(* Logix 5000 project; controller NWGG 1756-L72 rev 35.12; software revision 35.00; part 7 of 19 *)
(* tags used below, declared in another part *)
   _11_BINDICA : ALIAS FOR B15[11].0;
   _11_BINDICA1 : ALIAS FOR B15[11].1;
   _11_GATE_PO : ALIAS FOR I16[0];
   _11_GATE_PO1 : ALIAS FOR N14[11];
   _12_BINDICA : ALIAS FOR B15[12].0;
   _12_BINDICA1 : ALIAS FOR B15[12].1;
   _12_GATE_PO : ALIAS FOR I16[1];
   _12_GATE_PO1 : ALIAS FOR N14[12];
   _13_BINDICA : ALIAS FOR B15[13].0;
   _13_BINDICA1 : ALIAS FOR B15[13].1;
   _13_GATE_PO : ALIAS FOR I16[2];
   _13_GATE_PO1 : ALIAS FOR N14[13];
   _14_BINDICA : ALIAS FOR B15[14].0;
   _14_BINDICA1 : ALIAS FOR B15[14].1;
   _14_GATE_PO : ALIAS FOR I16[3];
   _14_GATE_PO1 : ALIAS FOR N14[14];
   _15_BINDICA : ALIAS FOR B15[15].0;
   _15_BINDICA1 : ALIAS FOR B15[15].1;
   _15_GATE_PO : ALIAS FOR I16[4];
   _15_GATE_PO1 : ALIAS FOR N14[15];
   _16_BINDICA : ALIAS FOR B15[16].0;
   _16_BINDICA1 : ALIAS FOR B15[16].1;
   _16_GATE_PO : ALIAS FOR I16[5];
   _16_GATE_PO1 : ALIAS FOR N14[16];
   _17_BINDICA : ALIAS FOR B15[17].0;
   _17_BINDICA1 : ALIAS FOR B15[17].1;
   _17_GATE_PO : ALIAS FOR I16[6];
   _17_GATE_PO1 : ALIAS FOR N14[17];
   _21_BINDICA : ALIAS FOR B15[21].0;
   _21_BINDICA1 : ALIAS FOR B15[21].1;
   _21_GATE_PO : ALIAS FOR I16[7];
   _21_GATE_PO1 : ALIAS FOR N14[21];
   _22_BINDICA : ALIAS FOR B15[22].0;
   _22_BINDICA1 : ALIAS FOR B15[22].1;
   _22_GATE_PO : ALIAS FOR I17[0];
   _22_GATE_PO1 : ALIAS FOR N14[22];
   _23_BINDICA : ALIAS FOR B15[23].0;
   _23_BINDICA1 : ALIAS FOR B15[23].1;
   _23_GATE_PO : ALIAS FOR I17[1];
   _23_GATE_PO1 : ALIAS FOR N14[23];
   _24_BINDICA : ALIAS FOR B15[24].0;
   _24_BINDICA1 : ALIAS FOR B15[24].1;
   _24_GATE_PO : ALIAS FOR I17[2];
   _24_GATE_PO1 : ALIAS FOR N14[24];
   _25_BINDICA : ALIAS FOR B15[25].0;
   _25_BINDICA1 : ALIAS FOR B15[25].1;
   _25_GATE_PO : ALIAS FOR I17[3];
   _25_GATE_PO1 : ALIAS FOR N14[25];
   _26_BINDICA : ALIAS FOR B15[26].0;
   _26_BINDICA1 : ALIAS FOR B15[26].1;
   _26_GATE_PO : ALIAS FOR I17[4];
   _26_GATE_PO1 : ALIAS FOR N14[26];
   _41_GATE_PO : ALIAS FOR I18[0];
   _41_GATE_PO1 : ALIAS FOR N14[41];
   _42_GATE_PO : ALIAS FOR I18[1];
   _42_GATE_PO1 : ALIAS FOR N14[42];
   _700_AIR_GA : ALIAS FOR I8.3;
   _701_AIR_GA : ALIAS FOR I8.5;
   _708G_BIN_1 : ALIAS FOR O9.15;
   _709G_BIN_1 : ALIAS FOR O10.15;
   A_HOLD_REL : ALIAS FOR B3[1].5;
   A_STPB_AUT : ALIAS FOR B3[1].1;
   Analog : AI[160];
   CAL_K_FACT : ALIAS FOR F8[0];
   CAL_RESET : ALIAS FOR B15[50].0;
   CIMBRA_BIN : ALIAS FOR I25[3].10;
   CIMBRIA_BI : ALIAS FOR B15[30].0;
   CIMBRIA_BI1 : ALIAS FOR B15[30].1;
   CIMBRIA_HI : ALIAS FOR B15[30].2;
   CONC13_PUM : ALIAS FOR N7[83];
   CONC19_PUM : ALIAS FOR N7[89];
   CONC_13_NO : ALIAS FOR B21[8].15;
   CONC_19_NO : ALIAS FOR B21[9].15;
   I1_000_Bit00 : ALIAS FOR I1.0;
   I1_000_Bit01 : ALIAS FOR I1.1;
   I1_000_Bit03 : ALIAS FOR I1.3;
   I1_000_Bit04 : ALIAS FOR I1.4;
   I1_000_Bit06 : ALIAS FOR I1.6;
   I1_000_Bit07 : ALIAS FOR I1.7;
   I1_000_Bit09 : ALIAS FOR I1.9;
   I1_000_Bit10 : ALIAS FOR I1.10;
   I1_000_Bit12 : ALIAS FOR I1.12;
   I1_000_Bit13 : ALIAS FOR I1.13;
   I1_000_Bit15 : ALIAS FOR I1.15;
   I24_021_Bit00 : ALIAS FOR I24[21].0;
   I24_021_Bit01 : ALIAS FOR I24[21].1;
   I24_021_Bit02 : ALIAS FOR I24[21].2;
   I2_000_Bit00 : ALIAS FOR I2.0;
   I2_000_Bit03 : ALIAS FOR I2.3;
   I2_000_Bit06 : ALIAS FOR I2.6;
   I2_000_Bit09 : ALIAS FOR I2.9;
   I2_000_Bit12 : ALIAS FOR I2.12;
   I3_000_Bit00 : ALIAS FOR I3.0;
   I3_000_Bit03 : ALIAS FOR I3.3;
   I3_000_Bit06 : ALIAS FOR I3.6;
   I4_000_Bit09 : ALIAS FOR I4.9;
   I4_000_Bit10 : ALIAS FOR I4.10;
   I4_000_Bit11 : ALIAS FOR I4.11;
   I4_000_Bit12 : ALIAS FOR I4.12;
   I4_000_Bit13 : ALIAS FOR I4.13;
   I4_000_Bit14 : ALIAS FOR I4.14;
   I4_000_Bit15 : ALIAS FOR I4.15;
   K_FACTOR : ALIAS FOR N14[80];
   P1_ALARM_N : ALIAS FOR T4[81];
   P1_ALARM_N1 : ALIAS FOR T4[82];
   P1_NO_FLOW : ALIAS FOR B12[1].3;
   P1_SEC_SEL : ALIAS FOR B17[1].1;
   P2_ALARM_N : ALIAS FOR T4[83];
   P2_ALARM_N1 : ALIAS FOR T4[84];
   P2_NO_FLOW : ALIAS FOR B12[2].3;
   P2_SEC_SEL : ALIAS FOR B17[1].2;
   P3_ALARM_N : ALIAS FOR T4[85];
   P3_ALARM_N1 : ALIAS FOR T4[86];
   P3_NO_FLOW : ALIAS FOR B12[3].3;
   P3_SEC_SEL : ALIAS FOR B17[1].3;
   P4_SEC_SEL : ALIAS FOR B17[1].4;
   T11_CAL_CL : ALIAS FOR B15[51].3;
   T11_CAL_LA : ALIAS FOR B15[51].2;
   T11_CAL_OP : ALIAS FOR B15[51].4;
   T11_CAL_ST : ALIAS FOR B15[51].1;
   T11_CORREC : ALIAS FOR F8[2];
   T11_K_FACT : ALIAS FOR F8[1];
   T11_LOW_BI : ALIAS FOR B15[11].2;
   T11_NO_PAS : ALIAS FOR B17[11].2;
   T12_CAL_CL : ALIAS FOR B15[52].3;
   T12_CAL_LA : ALIAS FOR B15[52].2;
   T12_CAL_OP : ALIAS FOR B15[52].4;
   T12_CAL_ST : ALIAS FOR B15[52].1;
   T12_CORREC : ALIAS FOR F8[4];
   T12_K_FACT : ALIAS FOR F8[3];
   T12_LOW_BI : ALIAS FOR B15[12].2;
   T12_NO_PAS : ALIAS FOR B17[12].2;
   T13_CAL_CL : ALIAS FOR B15[53].3;
   T13_CAL_LA : ALIAS FOR B15[53].2;
   T13_CAL_OP : ALIAS FOR B15[53].4;
   T13_CAL_ST : ALIAS FOR B15[53].1;
   T13_CORREC : ALIAS FOR F8[6];
   T13_K_FACT : ALIAS FOR F8[5];
   T13_LOW_BI : ALIAS FOR B15[13].2;
   T13_NO_PAS : ALIAS FOR B17[13].2;
   T14_CAL_CL : ALIAS FOR B15[54].3;
   T14_CAL_LA : ALIAS FOR B15[54].2;
   T14_CAL_OP : ALIAS FOR B15[54].4;
   T14_CAL_ST : ALIAS FOR B15[54].1;
   T14_CORREC : ALIAS FOR F8[8];
   T14_K_FACT : ALIAS FOR F8[7];
   T14_LOW_BI : ALIAS FOR B15[14].2;
   T14_NO_PAS : ALIAS FOR B17[14].2;
   T15_CAL_CL : ALIAS FOR B15[55].3;
   T15_CAL_LA : ALIAS FOR B15[55].2;
   T15_CAL_OP : ALIAS FOR B15[55].4;
   T15_CAL_ST : ALIAS FOR B15[55].1;
   T15_CORREC : ALIAS FOR F8[10];
   T15_K_FACT : ALIAS FOR F8[9];
   T15_LOW_BI : ALIAS FOR B15[15].2;
   T15_NO_PAS : ALIAS FOR B17[15].2;
   T16_CAL_CL : ALIAS FOR B15[56].3;
   T16_CAL_LA : ALIAS FOR B15[56].2;
   T16_CAL_OP : ALIAS FOR B15[56].4;
   T16_CAL_ST : ALIAS FOR B15[56].1;
   T16_CORREC : ALIAS FOR F8[12];
   T16_K_FACT : ALIAS FOR F8[11];
   T16_LOW_BI : ALIAS FOR B15[16].2;
   T16_NO_PAS : ALIAS FOR B17[16].2;
   T17_CAL_CL : ALIAS FOR B15[57].3;
   T17_CAL_LA : ALIAS FOR B15[57].2;
   T17_CAL_OP : ALIAS FOR B15[57].4;
   T17_CAL_ST : ALIAS FOR B15[57].1;
   T17_CORREC : ALIAS FOR F8[14];
   T17_K_FACT : ALIAS FOR F8[13];
   T17_LOW_BI : ALIAS FOR B15[17].2;
   T17_NO_PAS : ALIAS FOR B17[17].2;
   T21_CAL_CL : ALIAS FOR B15[61].3;
   T21_CAL_LA : ALIAS FOR B15[61].2;
   T21_CAL_OP : ALIAS FOR B15[61].4;
   T21_CAL_ST : ALIAS FOR B15[61].1;
   T21_CORREC : ALIAS FOR F8[16];
   T21_K_FACT : ALIAS FOR F8[15];
   T21_LOW_BI : ALIAS FOR B15[21].2;
   T21_NO_PAS : ALIAS FOR B17[21].2;
   T22_CAL_CL : ALIAS FOR B15[62].3;
   T22_CAL_LA : ALIAS FOR B15[62].2;
   T22_CAL_OP : ALIAS FOR B15[62].4;
   T22_CAL_ST : ALIAS FOR B15[62].1;
   T22_CORREC : ALIAS FOR F8[18];
   T22_K_FACT : ALIAS FOR F8[17];
   T22_LOW_BI : ALIAS FOR B15[22].2;
   T22_NO_PAS : ALIAS FOR B17[22].2;
   T23_CAL_CL : ALIAS FOR B15[63].3;
   T23_CAL_LA : ALIAS FOR B15[63].2;
   T23_CAL_OP : ALIAS FOR B15[63].4;
   T23_CAL_ST : ALIAS FOR B15[63].1;
   T23_CORREC : ALIAS FOR F8[20];
   T23_K_FACT : ALIAS FOR F8[19];
   T23_LOW_BI : ALIAS FOR B15[23].2;
   T23_NO_PAS : ALIAS FOR B17[23].2;
   T24_CAL_CL : ALIAS FOR B15[64].3;
   T24_CAL_LA : ALIAS FOR B15[64].2;
   T24_CAL_OP : ALIAS FOR B15[64].4;
   T24_CAL_ST : ALIAS FOR B15[64].1;
   T24_CORREC : ALIAS FOR F8[22];
   T24_K_FACT : ALIAS FOR F8[21];
   T24_LOW_BI : ALIAS FOR B15[24].2;
   T24_NO_PAS : ALIAS FOR B17[24].2;
   T25_CAL_CL : ALIAS FOR B15[65].3;
   T25_CAL_LA : ALIAS FOR B15[65].2;
   T25_CAL_OP : ALIAS FOR B15[65].4;
   T25_CAL_ST : ALIAS FOR B15[65].1;
   T25_CORREC : ALIAS FOR F8[24];
   T25_K_FACT : ALIAS FOR F8[23];
   T25_LOW_BI : ALIAS FOR B15[25].2;
   T25_NO_PAS : ALIAS FOR B17[25].2;
   T26_CAL_CL : ALIAS FOR B15[66].3;
   T26_CAL_LA : ALIAS FOR B15[66].2;
   T26_CAL_OP : ALIAS FOR B15[66].4;
   T26_CAL_ST : ALIAS FOR B15[66].1;
   T26_CORREC : ALIAS FOR F8[26];
   T26_K_FACT : ALIAS FOR F8[25];
   T26_LOW_BI : ALIAS FOR B15[26].2;
   T26_NO_PAS : ALIAS FOR B17[26].2;
   TK11_PUMP : ALIAS FOR N7[70];
   TK12_PUMP : ALIAS FOR N7[71];
   TK13_PUMP : ALIAS FOR N7[72];
   TK14_PUMP : ALIAS FOR N7[73];
   TK15_PUMP : ALIAS FOR N7[74];
   TK16_PUMP : ALIAS FOR N7[75];
   TK17_PUMP : ALIAS FOR N7[76];
   TK21_PUMP : ALIAS FOR N7[77];
   TK22_PUMP : ALIAS FOR N7[78];
   TK23_PUMP : ALIAS FOR N7[79];
   TK24_PUMP : ALIAS FOR N7[80];
   TK25_PUMP : ALIAS FOR N7[81];
   TK26_PUMP : ALIAS FOR N7[82];
(* _2_MAIN, continued *)

ROUTINE _37_BINDICATOR   (* ladder *)
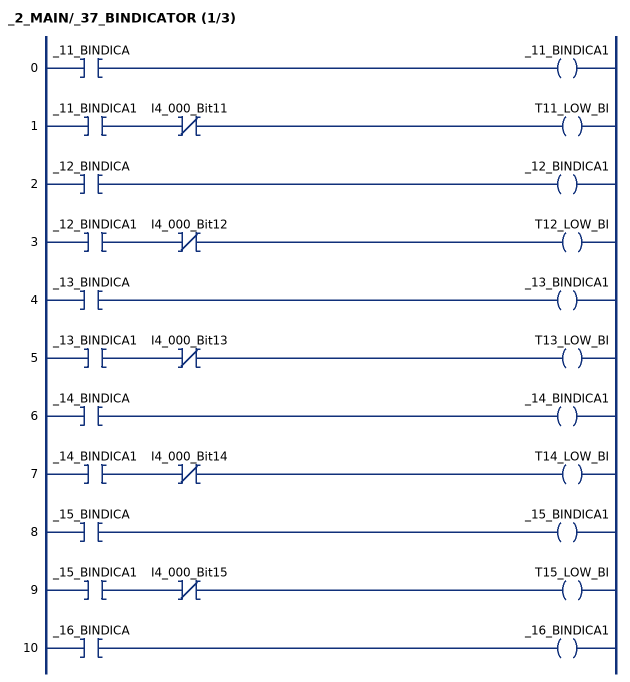
   0: XIC(_11_BINDICA)OTE(_11_BINDICA1);
   1: XIC(_11_BINDICA1)XIO(I4_000_Bit11)OTE(T11_LOW_BI);
   2: XIC(_12_BINDICA)OTE(_12_BINDICA1);
   3: XIC(_12_BINDICA1)XIO(I4_000_Bit12)OTE(T12_LOW_BI);
   4: XIC(_13_BINDICA)OTE(_13_BINDICA1);
   5: XIC(_13_BINDICA1)XIO(I4_000_Bit13)OTE(T13_LOW_BI);
   6: XIC(_14_BINDICA)OTE(_14_BINDICA1);
   7: XIC(_14_BINDICA1)XIO(I4_000_Bit14)OTE(T14_LOW_BI);
   8: XIC(_15_BINDICA)OTE(_15_BINDICA1);
   9: XIC(_15_BINDICA1)XIO(I4_000_Bit15)OTE(T15_LOW_BI);
   10: XIC(_16_BINDICA)OTE(_16_BINDICA1);
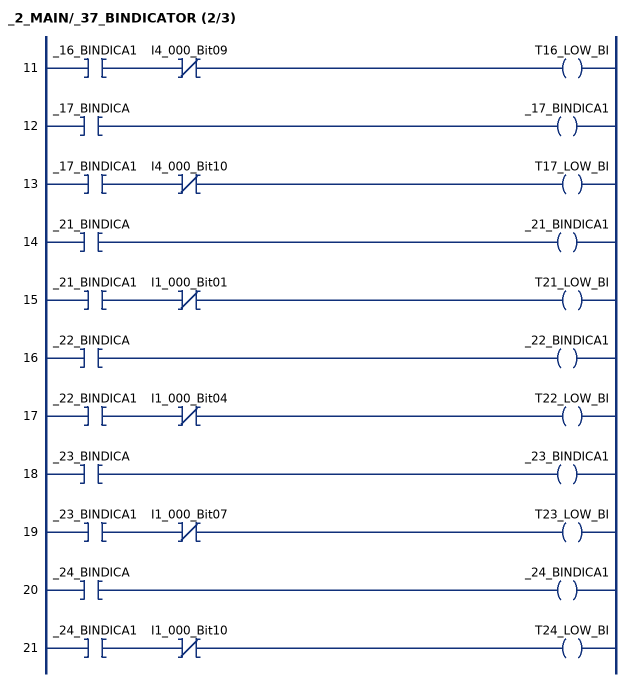
   11: XIC(_16_BINDICA1)XIO(I4_000_Bit09)OTE(T16_LOW_BI);
   12: XIC(_17_BINDICA)OTE(_17_BINDICA1);
   13: XIC(_17_BINDICA1)XIO(I4_000_Bit10)OTE(T17_LOW_BI);
   14: XIC(_21_BINDICA)OTE(_21_BINDICA1);
   15: XIC(_21_BINDICA1)XIO(I1_000_Bit01)OTE(T21_LOW_BI);
   16: XIC(_22_BINDICA)OTE(_22_BINDICA1);
   17: XIC(_22_BINDICA1)XIO(I1_000_Bit04)OTE(T22_LOW_BI);
   18: XIC(_23_BINDICA)OTE(_23_BINDICA1);
   19: XIC(_23_BINDICA1)XIO(I1_000_Bit07)OTE(T23_LOW_BI);
   20: XIC(_24_BINDICA)OTE(_24_BINDICA1);
   21: XIC(_24_BINDICA1)XIO(I1_000_Bit10)OTE(T24_LOW_BI);
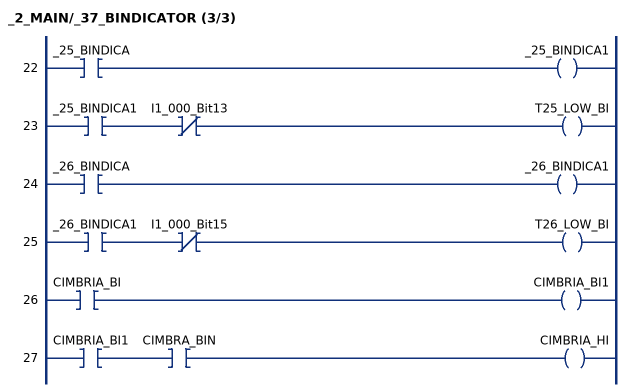
   22: XIC(_25_BINDICA)OTE(_25_BINDICA1);
   23: XIC(_25_BINDICA1)XIO(I1_000_Bit13)OTE(T25_LOW_BI);
   24: XIC(_26_BINDICA)OTE(_26_BINDICA1);
   25: XIC(_26_BINDICA1)XIO(I1_000_Bit15)OTE(T26_LOW_BI);
   26: XIC(CIMBRIA_BI)OTE(CIMBRIA_BI1);
   27: XIC(CIMBRIA_BI1)XIC(CIMBRA_BIN)OTE(CIMBRIA_HI);
END_ROUTINE

ROUTINE _38_GATE_ADJST   (* ladder *)
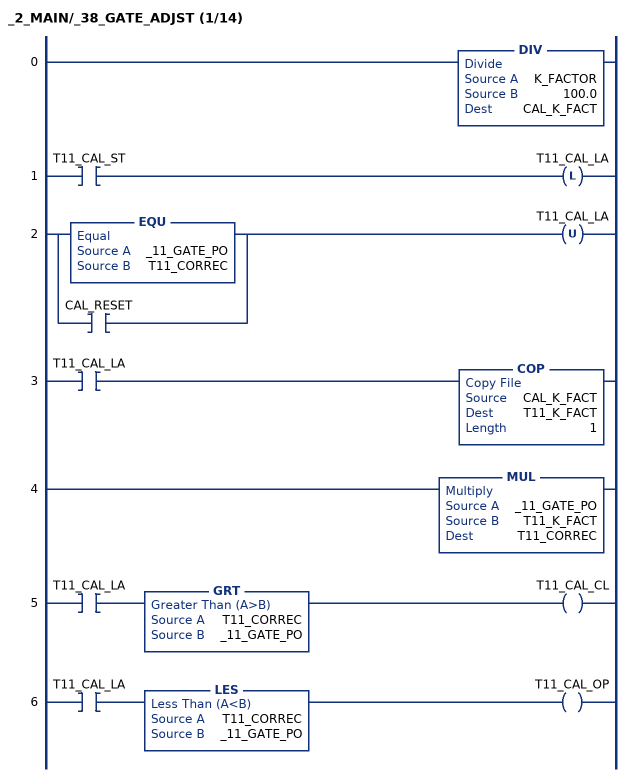
   0: DIV(K_FACTOR,100.0,CAL_K_FACT);
   1: XIC(T11_CAL_ST)OTL(T11_CAL_LA);
   2: [EQU(_11_GATE_PO,T11_CORREC) ,XIC(CAL_RESET) ]OTU(T11_CAL_LA);
   3: XIC(T11_CAL_LA)COP(CAL_K_FACT,T11_K_FACT,1);
   4: MUL(_11_GATE_PO,T11_K_FACT,T11_CORREC);
   5: XIC(T11_CAL_LA)GRT(T11_CORREC,_11_GATE_PO)OTE(T11_CAL_CL);
   6: XIC(T11_CAL_LA)LES(T11_CORREC,_11_GATE_PO)OTE(T11_CAL_OP);
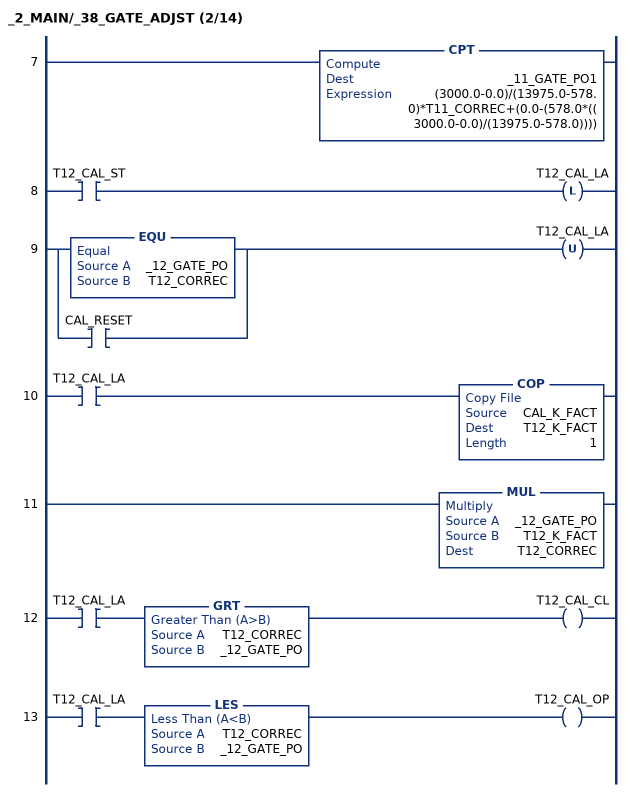
   7: CPT(_11_GATE_PO1,(3000.0-0.0)/(13975.0-578.0)*T11_CORREC+(0.0-(578.0*((3000.0-0.0)/(13975.0-578.0)))));
   8: XIC(T12_CAL_ST)OTL(T12_CAL_LA);
   9: [EQU(_12_GATE_PO,T12_CORREC) ,XIC(CAL_RESET) ]OTU(T12_CAL_LA);
   10: XIC(T12_CAL_LA)COP(CAL_K_FACT,T12_K_FACT,1);
   11: MUL(_12_GATE_PO,T12_K_FACT,T12_CORREC);
   12: XIC(T12_CAL_LA)GRT(T12_CORREC,_12_GATE_PO)OTE(T12_CAL_CL);
   13: XIC(T12_CAL_LA)LES(T12_CORREC,_12_GATE_PO)OTE(T12_CAL_OP);
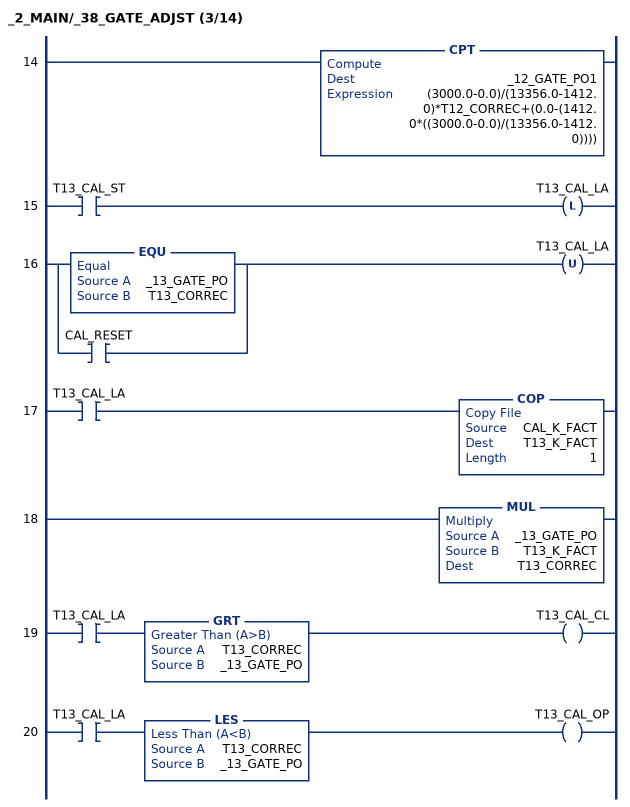
   14: CPT(_12_GATE_PO1,(3000.0-0.0)/(13356.0-1412.0)*T12_CORREC+(0.0-(1412.0*((3000.0-0.0)/(13356.0-1412.0)))));
   15: XIC(T13_CAL_ST)OTL(T13_CAL_LA);
   16: [EQU(_13_GATE_PO,T13_CORREC) ,XIC(CAL_RESET) ]OTU(T13_CAL_LA);
   17: XIC(T13_CAL_LA)COP(CAL_K_FACT,T13_K_FACT,1);
   18: MUL(_13_GATE_PO,T13_K_FACT,T13_CORREC);
   19: XIC(T13_CAL_LA)GRT(T13_CORREC,_13_GATE_PO)OTE(T13_CAL_CL);
   20: XIC(T13_CAL_LA)LES(T13_CORREC,_13_GATE_PO)OTE(T13_CAL_OP);
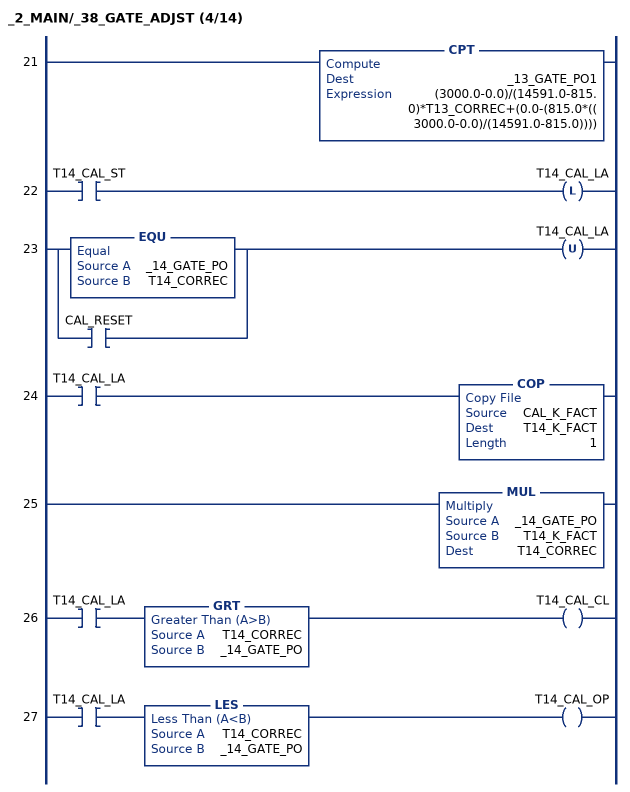
   21: CPT(_13_GATE_PO1,(3000.0-0.0)/(14591.0-815.0)*T13_CORREC+(0.0-(815.0*((3000.0-0.0)/(14591.0-815.0)))));
   22: XIC(T14_CAL_ST)OTL(T14_CAL_LA);
   23: [EQU(_14_GATE_PO,T14_CORREC) ,XIC(CAL_RESET) ]OTU(T14_CAL_LA);
   24: XIC(T14_CAL_LA)COP(CAL_K_FACT,T14_K_FACT,1);
   25: MUL(_14_GATE_PO,T14_K_FACT,T14_CORREC);
   26: XIC(T14_CAL_LA)GRT(T14_CORREC,_14_GATE_PO)OTE(T14_CAL_CL);
   27: XIC(T14_CAL_LA)LES(T14_CORREC,_14_GATE_PO)OTE(T14_CAL_OP);
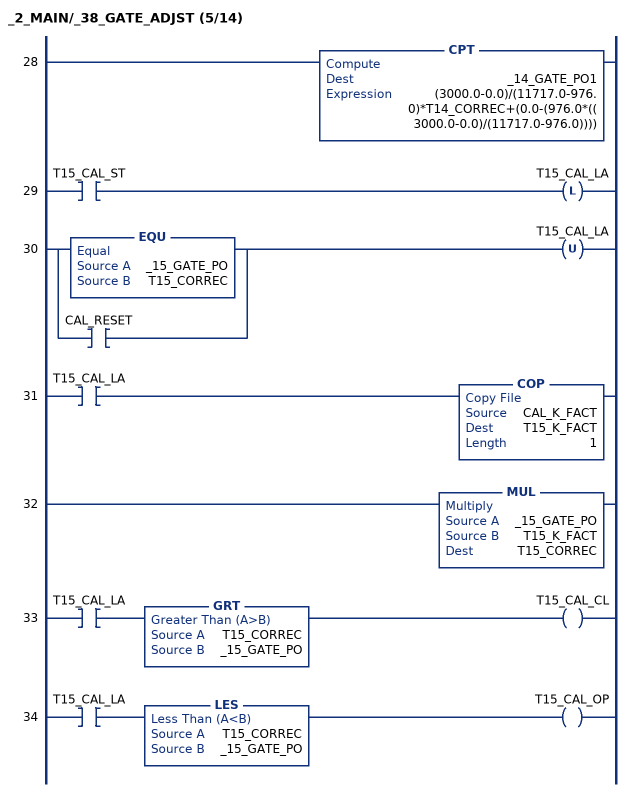
   28: CPT(_14_GATE_PO1,(3000.0-0.0)/(11717.0-976.0)*T14_CORREC+(0.0-(976.0*((3000.0-0.0)/(11717.0-976.0)))));
   29: XIC(T15_CAL_ST)OTL(T15_CAL_LA);
   30: [EQU(_15_GATE_PO,T15_CORREC) ,XIC(CAL_RESET) ]OTU(T15_CAL_LA);
   31: XIC(T15_CAL_LA)COP(CAL_K_FACT,T15_K_FACT,1);
   32: MUL(_15_GATE_PO,T15_K_FACT,T15_CORREC);
   33: XIC(T15_CAL_LA)GRT(T15_CORREC,_15_GATE_PO)OTE(T15_CAL_CL);
   34: XIC(T15_CAL_LA)LES(T15_CORREC,_15_GATE_PO)OTE(T15_CAL_OP);
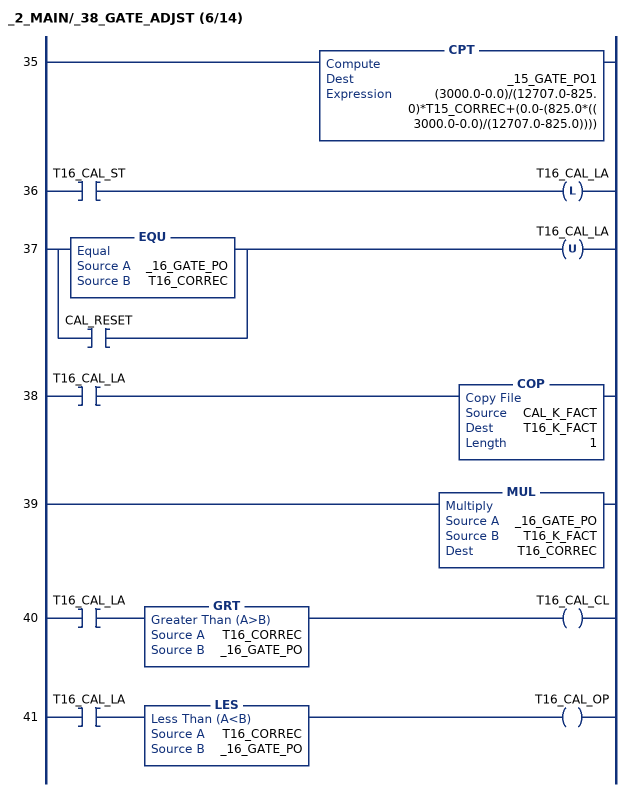
   35: CPT(_15_GATE_PO1,(3000.0-0.0)/(12707.0-825.0)*T15_CORREC+(0.0-(825.0*((3000.0-0.0)/(12707.0-825.0)))));
   36: XIC(T16_CAL_ST)OTL(T16_CAL_LA);
   37: [EQU(_16_GATE_PO,T16_CORREC) ,XIC(CAL_RESET) ]OTU(T16_CAL_LA);
   38: XIC(T16_CAL_LA)COP(CAL_K_FACT,T16_K_FACT,1);
   39: MUL(_16_GATE_PO,T16_K_FACT,T16_CORREC);
   40: XIC(T16_CAL_LA)GRT(T16_CORREC,_16_GATE_PO)OTE(T16_CAL_CL);
   41: XIC(T16_CAL_LA)LES(T16_CORREC,_16_GATE_PO)OTE(T16_CAL_OP);
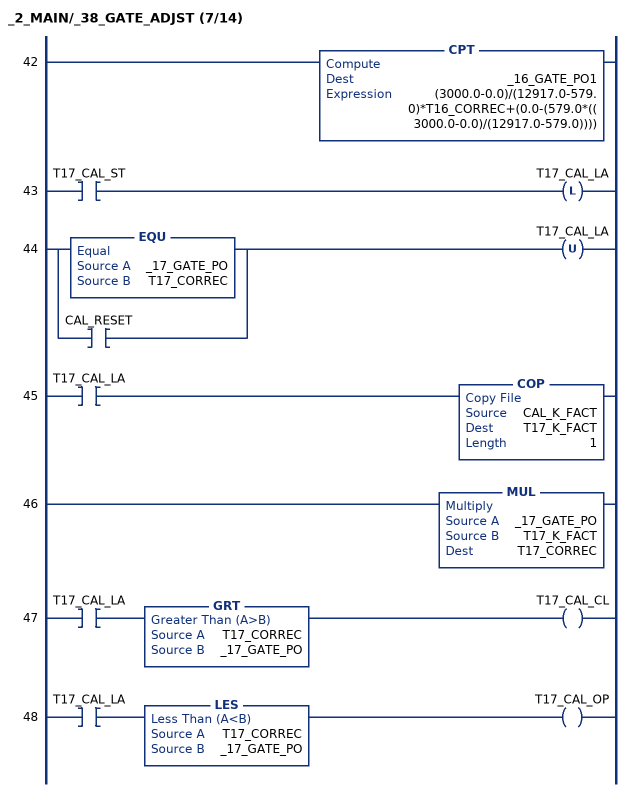
   42: CPT(_16_GATE_PO1,(3000.0-0.0)/(12917.0-579.0)*T16_CORREC+(0.0-(579.0*((3000.0-0.0)/(12917.0-579.0)))));
   43: XIC(T17_CAL_ST)OTL(T17_CAL_LA);
   44: [EQU(_17_GATE_PO,T17_CORREC) ,XIC(CAL_RESET) ]OTU(T17_CAL_LA);
   45: XIC(T17_CAL_LA)COP(CAL_K_FACT,T17_K_FACT,1);
   46: MUL(_17_GATE_PO,T17_K_FACT,T17_CORREC);
   47: XIC(T17_CAL_LA)GRT(T17_CORREC,_17_GATE_PO)OTE(T17_CAL_CL);
   48: XIC(T17_CAL_LA)LES(T17_CORREC,_17_GATE_PO)OTE(T17_CAL_OP);
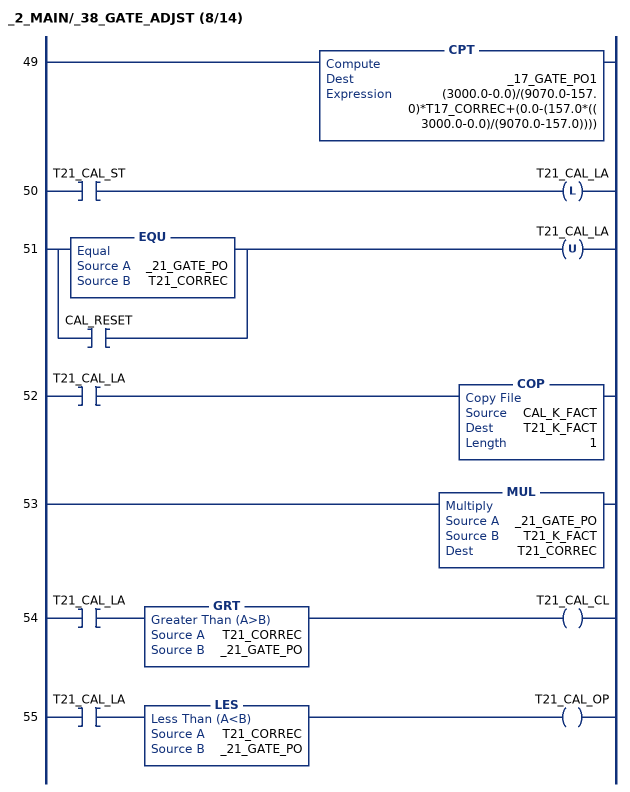
   49: CPT(_17_GATE_PO1,(3000.0-0.0)/(9070.0-157.0)*T17_CORREC+(0.0-(157.0*((3000.0-0.0)/(9070.0-157.0)))));
   50: XIC(T21_CAL_ST)OTL(T21_CAL_LA);
   51: [EQU(_21_GATE_PO,T21_CORREC) ,XIC(CAL_RESET) ]OTU(T21_CAL_LA);
   52: XIC(T21_CAL_LA)COP(CAL_K_FACT,T21_K_FACT,1);
   53: MUL(_21_GATE_PO,T21_K_FACT,T21_CORREC);
   54: XIC(T21_CAL_LA)GRT(T21_CORREC,_21_GATE_PO)OTE(T21_CAL_CL);
   55: XIC(T21_CAL_LA)LES(T21_CORREC,_21_GATE_PO)OTE(T21_CAL_OP);
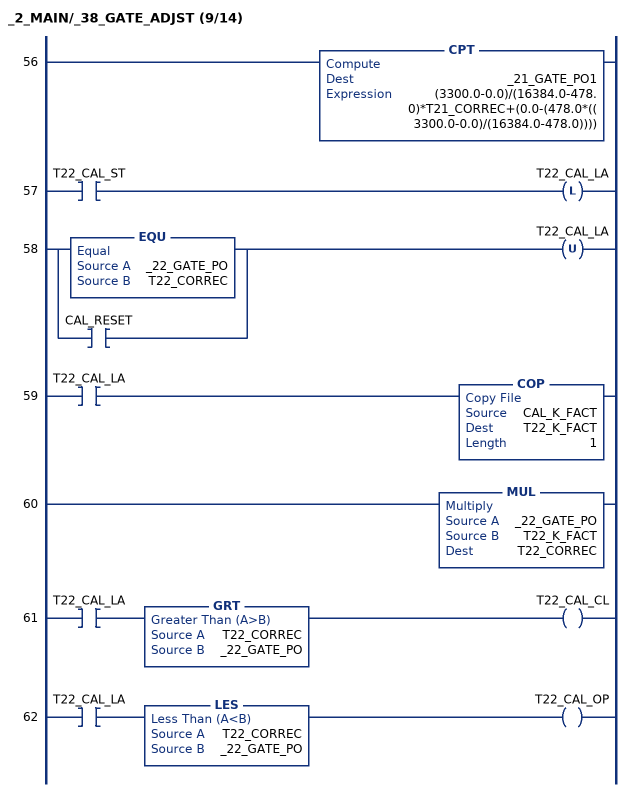
   56: CPT(_21_GATE_PO1,(3300.0-0.0)/(16384.0-478.0)*T21_CORREC+(0.0-(478.0*((3300.0-0.0)/(16384.0-478.0)))));
   57: XIC(T22_CAL_ST)OTL(T22_CAL_LA);
   58: [EQU(_22_GATE_PO,T22_CORREC) ,XIC(CAL_RESET) ]OTU(T22_CAL_LA);
   59: XIC(T22_CAL_LA)COP(CAL_K_FACT,T22_K_FACT,1);
   60: MUL(_22_GATE_PO,T22_K_FACT,T22_CORREC);
   61: XIC(T22_CAL_LA)GRT(T22_CORREC,_22_GATE_PO)OTE(T22_CAL_CL);
   62: XIC(T22_CAL_LA)LES(T22_CORREC,_22_GATE_PO)OTE(T22_CAL_OP);
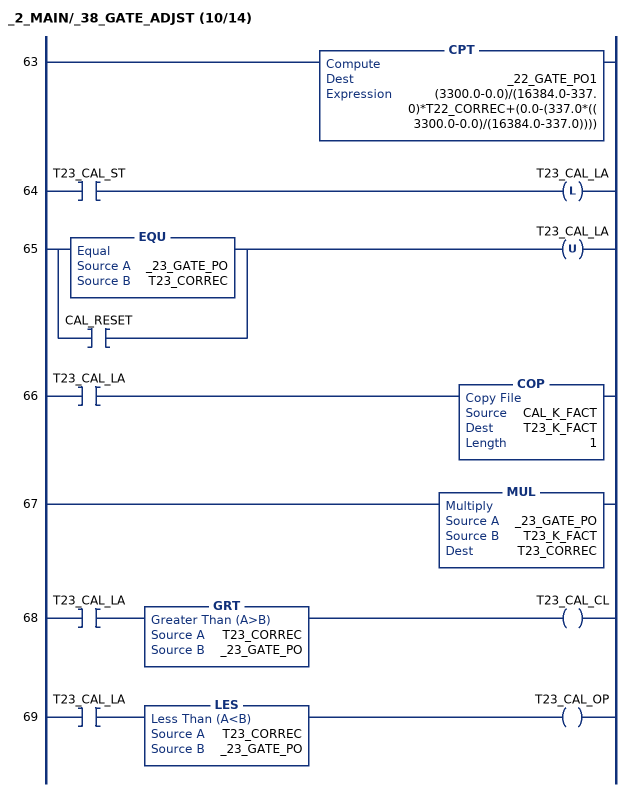
   63: CPT(_22_GATE_PO1,(3300.0-0.0)/(16384.0-337.0)*T22_CORREC+(0.0-(337.0*((3300.0-0.0)/(16384.0-337.0)))));
   64: XIC(T23_CAL_ST)OTL(T23_CAL_LA);
   65: [EQU(_23_GATE_PO,T23_CORREC) ,XIC(CAL_RESET) ]OTU(T23_CAL_LA);
   66: XIC(T23_CAL_LA)COP(CAL_K_FACT,T23_K_FACT,1);
   67: MUL(_23_GATE_PO,T23_K_FACT,T23_CORREC);
   68: XIC(T23_CAL_LA)GRT(T23_CORREC,_23_GATE_PO)OTE(T23_CAL_CL);
   69: XIC(T23_CAL_LA)LES(T23_CORREC,_23_GATE_PO)OTE(T23_CAL_OP);
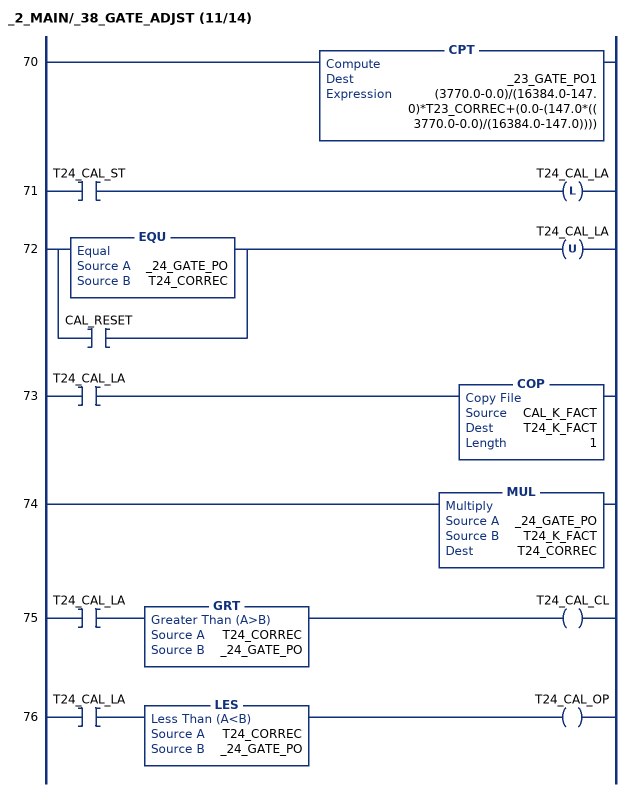
   70: CPT(_23_GATE_PO1,(3770.0-0.0)/(16384.0-147.0)*T23_CORREC+(0.0-(147.0*((3770.0-0.0)/(16384.0-147.0)))));
   71: XIC(T24_CAL_ST)OTL(T24_CAL_LA);
   72: [EQU(_24_GATE_PO,T24_CORREC) ,XIC(CAL_RESET) ]OTU(T24_CAL_LA);
   73: XIC(T24_CAL_LA)COP(CAL_K_FACT,T24_K_FACT,1);
   74: MUL(_24_GATE_PO,T24_K_FACT,T24_CORREC);
   75: XIC(T24_CAL_LA)GRT(T24_CORREC,_24_GATE_PO)OTE(T24_CAL_CL);
   76: XIC(T24_CAL_LA)LES(T24_CORREC,_24_GATE_PO)OTE(T24_CAL_OP);
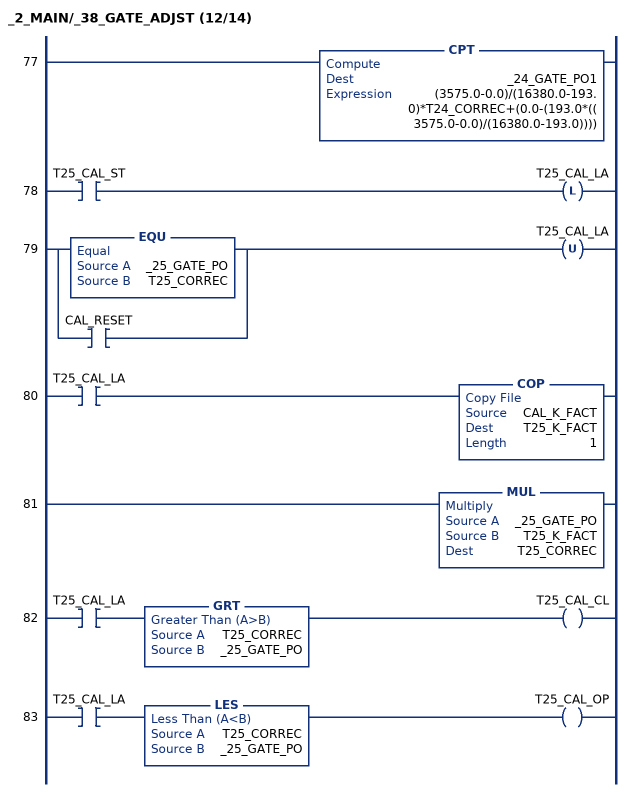
   77: CPT(_24_GATE_PO1,(3575.0-0.0)/(16380.0-193.0)*T24_CORREC+(0.0-(193.0*((3575.0-0.0)/(16380.0-193.0)))));
   78: XIC(T25_CAL_ST)OTL(T25_CAL_LA);
   79: [EQU(_25_GATE_PO,T25_CORREC) ,XIC(CAL_RESET) ]OTU(T25_CAL_LA);
   80: XIC(T25_CAL_LA)COP(CAL_K_FACT,T25_K_FACT,1);
   81: MUL(_25_GATE_PO,T25_K_FACT,T25_CORREC);
   82: XIC(T25_CAL_LA)GRT(T25_CORREC,_25_GATE_PO)OTE(T25_CAL_CL);
   83: XIC(T25_CAL_LA)LES(T25_CORREC,_25_GATE_PO)OTE(T25_CAL_OP);
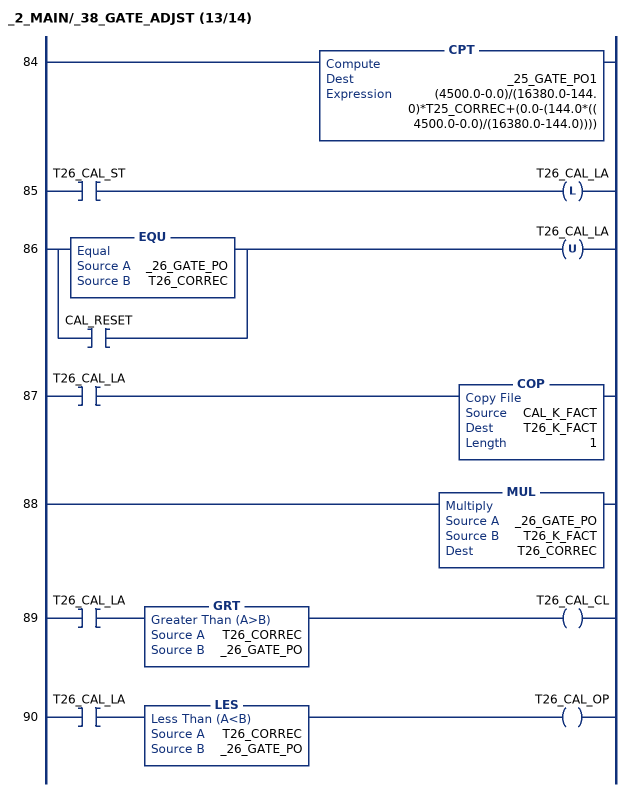
   84: CPT(_25_GATE_PO1,(4500.0-0.0)/(16380.0-144.0)*T25_CORREC+(0.0-(144.0*((4500.0-0.0)/(16380.0-144.0)))));
   85: XIC(T26_CAL_ST)OTL(T26_CAL_LA);
   86: [EQU(_26_GATE_PO,T26_CORREC) ,XIC(CAL_RESET) ]OTU(T26_CAL_LA);
   87: XIC(T26_CAL_LA)COP(CAL_K_FACT,T26_K_FACT,1);
   88: MUL(_26_GATE_PO,T26_K_FACT,T26_CORREC);
   89: XIC(T26_CAL_LA)GRT(T26_CORREC,_26_GATE_PO)OTE(T26_CAL_CL);
   90: XIC(T26_CAL_LA)LES(T26_CORREC,_26_GATE_PO)OTE(T26_CAL_OP);
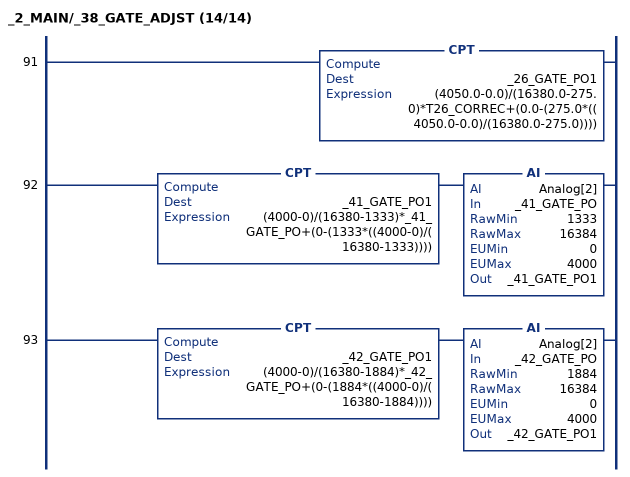
   91: CPT(_26_GATE_PO1,(4050.0-0.0)/(16380.0-275.0)*T26_CORREC+(0.0-(275.0*((4050.0-0.0)/(16380.0-275.0)))));
   92: CPT(_41_GATE_PO1,(4000-0)/(16380-1333)*_41_GATE_PO+(0-(1333*((4000-0)/(16380-1333)))))AI(Analog[2],_41_GATE_PO,1333,16384,0,4000,_41_GATE_PO1);
   93: CPT(_42_GATE_PO1,(4000-0)/(16380-1884)*_42_GATE_PO+(0-(1884*((4000-0)/(16380-1884)))))AI(Analog[2],_42_GATE_PO,1884,16384,0,4000,_42_GATE_PO1);
END_ROUTINE

ROUTINE _39_PUMP_SECUR   (* ladder *)
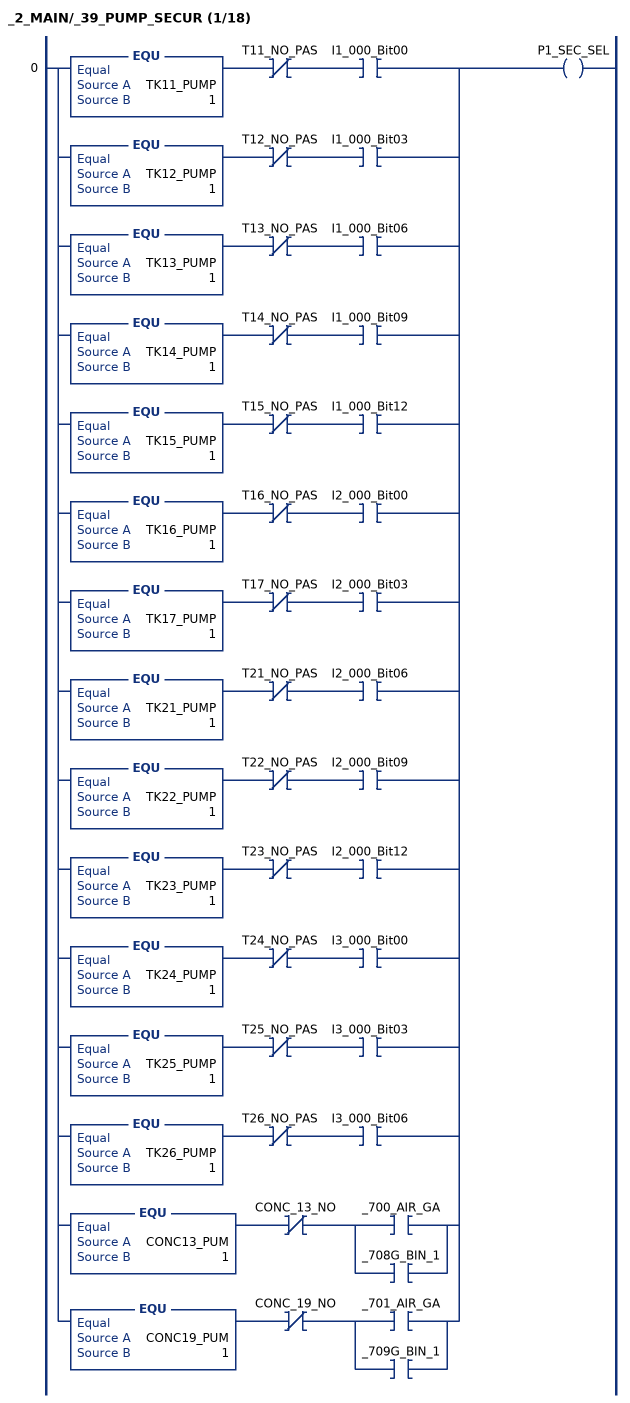
   0: [EQU(TK11_PUMP,1) XIO(T11_NO_PAS) XIC(I1_000_Bit00) ,EQU(TK12_PUMP,1) XIO(T12_NO_PAS) XIC(I1_000_Bit03) ,EQU(TK13_PUMP,1) XIO(T13_NO_PAS) XIC(I1_000_Bit06) ,EQU(TK14_PUMP,1) XIO(T14_NO_PAS) XIC(I1_000_Bit09) ,EQU(TK15_PUMP,1) XIO(T15_NO_PAS) XIC(I1_000_Bit12) ,EQU(TK16_PUMP,1) XIO(T16_NO_PAS) XIC(I2_000_Bit00) ,EQU(TK17_PUMP,1) XIO(T17_NO_PAS) XIC(I2_000_Bit03) ,EQU(TK21_PUMP,1) XIO(T21_NO_PAS) XIC(I2_000_Bit06) ,EQU(TK22_PUMP,1) XIO(T22_NO_PAS) XIC(I2_000_Bit09) ,EQU(TK23_PUMP,1) XIO(T23_NO_PAS) XIC(I2_000_Bit12) ,EQU(TK24_PUMP,1) XIO(T24_NO_PAS) XIC(I3_000_Bit00) ,EQU(TK25_PUMP,1) XIO(T25_NO_PAS) XIC(I3_000_Bit03) ,EQU(TK26_PUMP,1) XIO(T26_NO_PAS) XIC(I3_000_Bit06) ,EQU(CONC13_PUM,1) XIO(CONC_13_NO) [XIC(_700_AIR_GA) ,XIC(_708G_BIN_1) ] ,EQU(CONC19_PUM,1) XIO(CONC_19_NO) [XIC(_701_AIR_GA) ,XIC(_709G_BIN_1) ] ]OTE(P1_SEC_SEL);
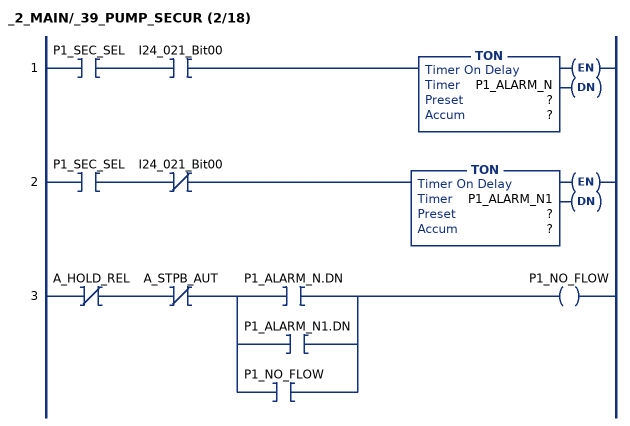
   1: XIC(P1_SEC_SEL)XIC(I24_021_Bit00)TON(P1_ALARM_N,?,?);
   2: XIC(P1_SEC_SEL)XIO(I24_021_Bit00)TON(P1_ALARM_N1,?,?);
   3: XIO(A_HOLD_REL)XIO(A_STPB_AUT)[XIC(P1_ALARM_N.DN) ,XIC(P1_ALARM_N1.DN) ,XIC(P1_NO_FLOW) ]OTE(P1_NO_FLOW);
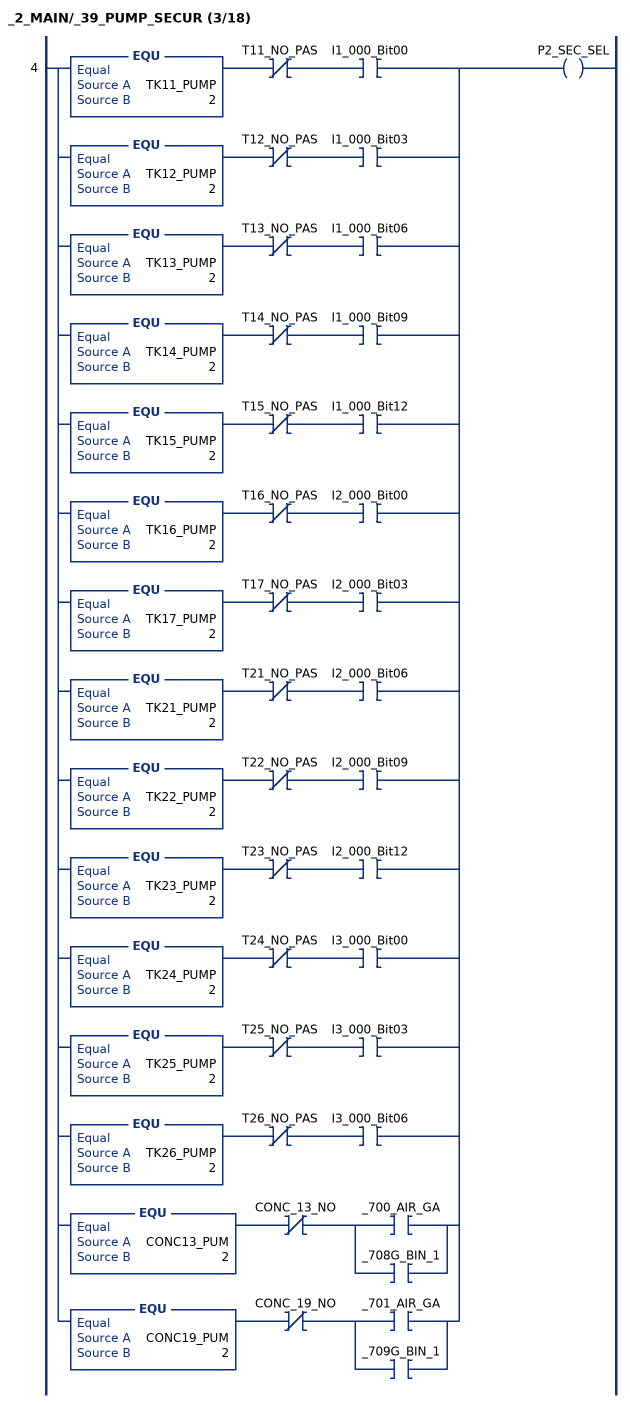
   4: [EQU(TK11_PUMP,2) XIO(T11_NO_PAS) XIC(I1_000_Bit00) ,EQU(TK12_PUMP,2) XIO(T12_NO_PAS) XIC(I1_000_Bit03) ,EQU(TK13_PUMP,2) XIO(T13_NO_PAS) XIC(I1_000_Bit06) ,EQU(TK14_PUMP,2) XIO(T14_NO_PAS) XIC(I1_000_Bit09) ,EQU(TK15_PUMP,2) XIO(T15_NO_PAS) XIC(I1_000_Bit12) ,EQU(TK16_PUMP,2) XIO(T16_NO_PAS) XIC(I2_000_Bit00) ,EQU(TK17_PUMP,2) XIO(T17_NO_PAS) XIC(I2_000_Bit03) ,EQU(TK21_PUMP,2) XIO(T21_NO_PAS) XIC(I2_000_Bit06) ,EQU(TK22_PUMP,2) XIO(T22_NO_PAS) XIC(I2_000_Bit09) ,EQU(TK23_PUMP,2) XIO(T23_NO_PAS) XIC(I2_000_Bit12) ,EQU(TK24_PUMP,2) XIO(T24_NO_PAS) XIC(I3_000_Bit00) ,EQU(TK25_PUMP,2) XIO(T25_NO_PAS) XIC(I3_000_Bit03) ,EQU(TK26_PUMP,2) XIO(T26_NO_PAS) XIC(I3_000_Bit06) ,EQU(CONC13_PUM,2) XIO(CONC_13_NO) [XIC(_700_AIR_GA) ,XIC(_708G_BIN_1) ] ,EQU(CONC19_PUM,2) XIO(CONC_19_NO) [XIC(_701_AIR_GA) ,XIC(_709G_BIN_1) ] ]OTE(P2_SEC_SEL);
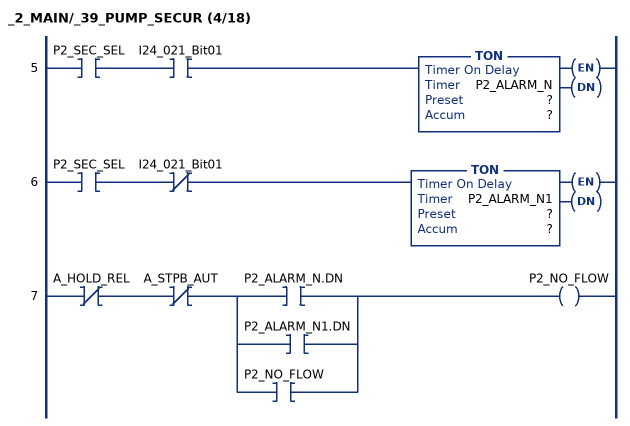
   5: XIC(P2_SEC_SEL)XIC(I24_021_Bit01)TON(P2_ALARM_N,?,?);
   6: XIC(P2_SEC_SEL)XIO(I24_021_Bit01)TON(P2_ALARM_N1,?,?);
   7: XIO(A_HOLD_REL)XIO(A_STPB_AUT)[XIC(P2_ALARM_N.DN) ,XIC(P2_ALARM_N1.DN) ,XIC(P2_NO_FLOW) ]OTE(P2_NO_FLOW);
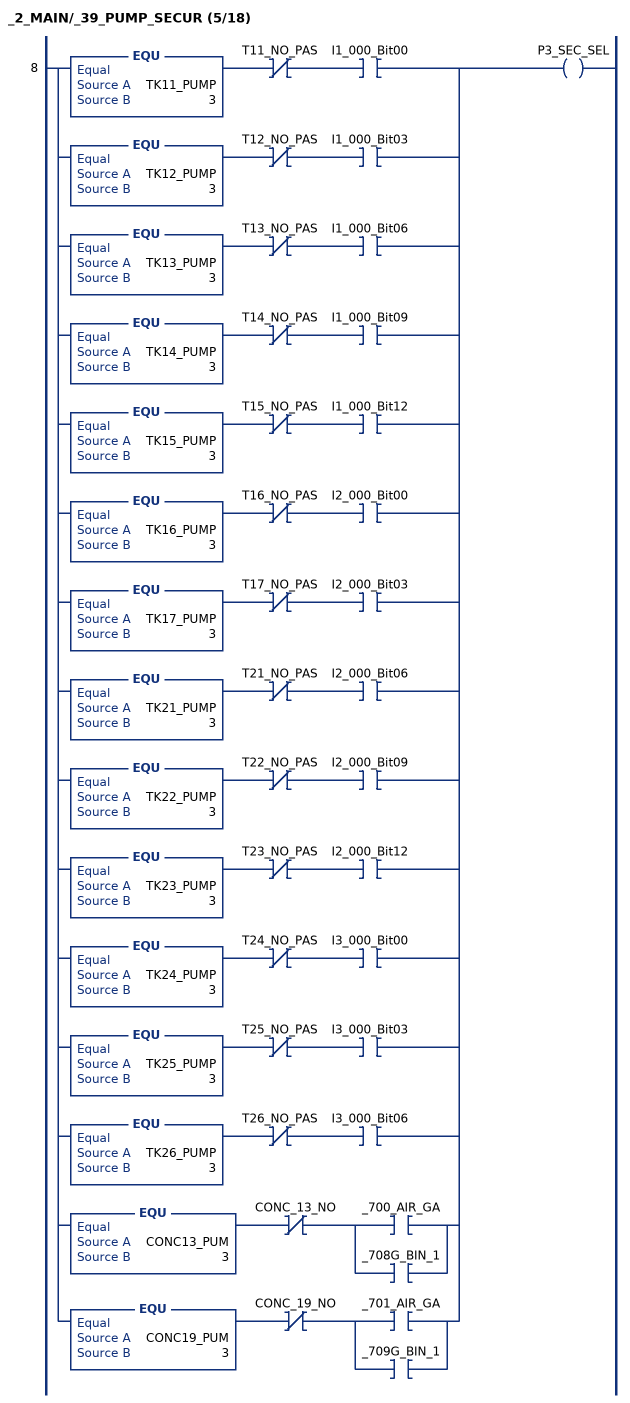
   8: [EQU(TK11_PUMP,3) XIO(T11_NO_PAS) XIC(I1_000_Bit00) ,EQU(TK12_PUMP,3) XIO(T12_NO_PAS) XIC(I1_000_Bit03) ,EQU(TK13_PUMP,3) XIO(T13_NO_PAS) XIC(I1_000_Bit06) ,EQU(TK14_PUMP,3) XIO(T14_NO_PAS) XIC(I1_000_Bit09) ,EQU(TK15_PUMP,3) XIO(T15_NO_PAS) XIC(I1_000_Bit12) ,EQU(TK16_PUMP,3) XIO(T16_NO_PAS) XIC(I2_000_Bit00) ,EQU(TK17_PUMP,3) XIO(T17_NO_PAS) XIC(I2_000_Bit03) ,EQU(TK21_PUMP,3) XIO(T21_NO_PAS) XIC(I2_000_Bit06) ,EQU(TK22_PUMP,3) XIO(T22_NO_PAS) XIC(I2_000_Bit09) ,EQU(TK23_PUMP,3) XIO(T23_NO_PAS) XIC(I2_000_Bit12) ,EQU(TK24_PUMP,3) XIO(T24_NO_PAS) XIC(I3_000_Bit00) ,EQU(TK25_PUMP,3) XIO(T25_NO_PAS) XIC(I3_000_Bit03) ,EQU(TK26_PUMP,3) XIO(T26_NO_PAS) XIC(I3_000_Bit06) ,EQU(CONC13_PUM,3) XIO(CONC_13_NO) [XIC(_700_AIR_GA) ,XIC(_708G_BIN_1) ] ,EQU(CONC19_PUM,3) XIO(CONC_19_NO) [XIC(_701_AIR_GA) ,XIC(_709G_BIN_1) ] ]OTE(P3_SEC_SEL);
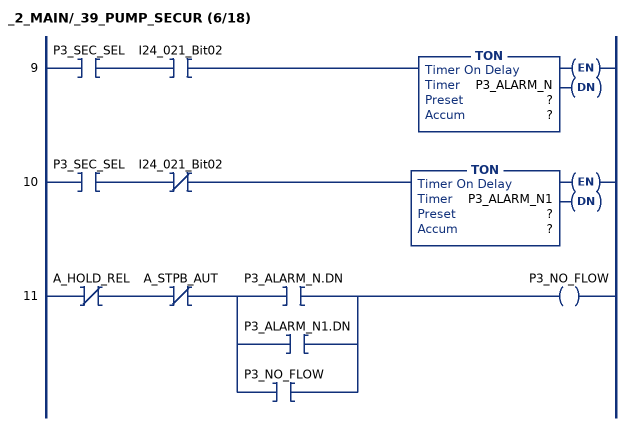
   9: XIC(P3_SEC_SEL)XIC(I24_021_Bit02)TON(P3_ALARM_N,?,?);
   10: XIC(P3_SEC_SEL)XIO(I24_021_Bit02)TON(P3_ALARM_N1,?,?);
   11: XIO(A_HOLD_REL)XIO(A_STPB_AUT)[XIC(P3_ALARM_N.DN) ,XIC(P3_ALARM_N1.DN) ,XIC(P3_NO_FLOW) ]OTE(P3_NO_FLOW);
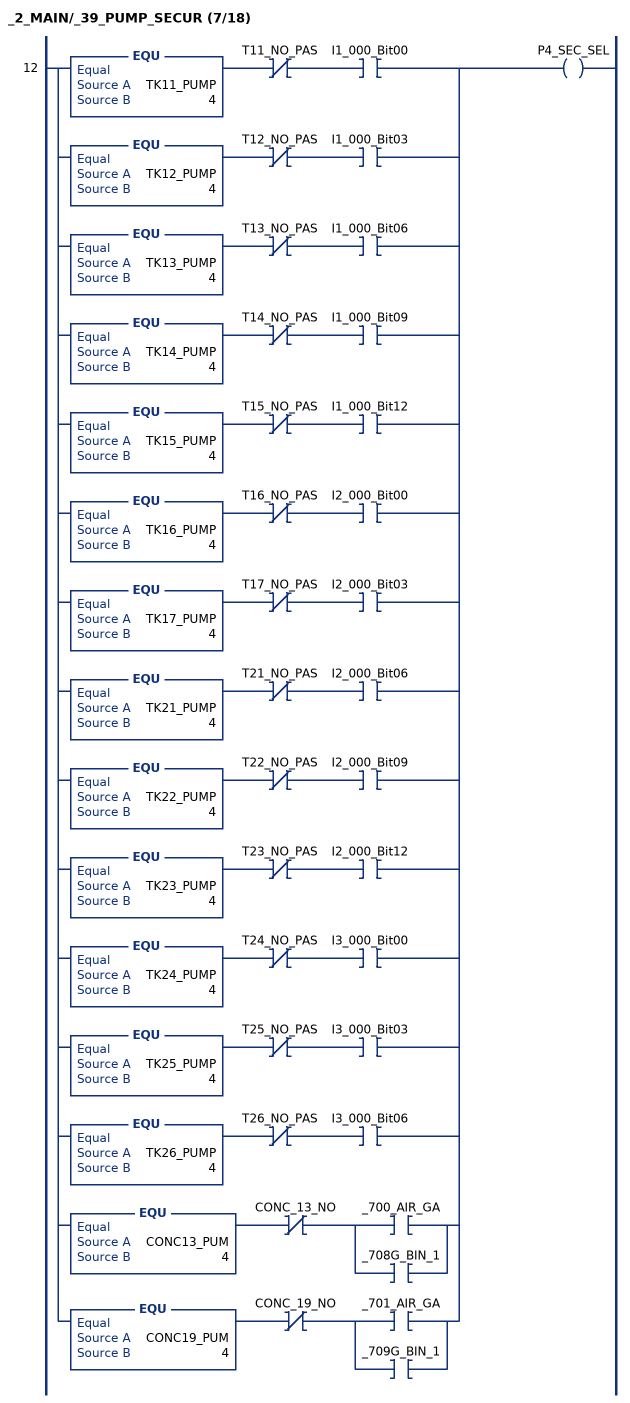
   12: [EQU(TK11_PUMP,4) XIO(T11_NO_PAS) XIC(I1_000_Bit00) ,EQU(TK12_PUMP,4) XIO(T12_NO_PAS) XIC(I1_000_Bit03) ,EQU(TK13_PUMP,4) XIO(T13_NO_PAS) XIC(I1_000_Bit06) ,EQU(TK14_PUMP,4) XIO(T14_NO_PAS) XIC(I1_000_Bit09) ,EQU(TK15_PUMP,4) XIO(T15_NO_PAS) XIC(I1_000_Bit12) ,EQU(TK16_PUMP,4) XIO(T16_NO_PAS) XIC(I2_000_Bit00) ,EQU(TK17_PUMP,4) XIO(T17_NO_PAS) XIC(I2_000_Bit03) ,EQU(TK21_PUMP,4) XIO(T21_NO_PAS) XIC(I2_000_Bit06) ,EQU(TK22_PUMP,4) XIO(T22_NO_PAS) XIC(I2_000_Bit09) ,EQU(TK23_PUMP,4) XIO(T23_NO_PAS) XIC(I2_000_Bit12) ,EQU(TK24_PUMP,4) XIO(T24_NO_PAS) XIC(I3_000_Bit00) ,EQU(TK25_PUMP,4) XIO(T25_NO_PAS) XIC(I3_000_Bit03) ,EQU(TK26_PUMP,4) XIO(T26_NO_PAS) XIC(I3_000_Bit06) ,EQU(CONC13_PUM,4) XIO(CONC_13_NO) [XIC(_700_AIR_GA) ,XIC(_708G_BIN_1) ] ,EQU(CONC19_PUM,4) XIO(CONC_19_NO) [XIC(_701_AIR_GA) ,XIC(_709G_BIN_1) ] ]OTE(P4_SEC_SEL);
